PROGRAM MAIN
VAR
END_VAR

ModbusMasterApplication;

END_PROGRAM

(* stored: Version 1.1.0.1, ProductVersion 3.1.4024.9
   POU MAIN: Id {af35dda5-7604-453c-8ab0-4b903fea5f9d}, SpecialFunc None *)
